Fanuc KAREL source: KT00636.KL

PROGRAM KT00636
%NOLOCKGROUP
VAR
  Y1: ARRAY[2] OF BYTE
  Y2: ARRAY[2] OF BYTE
  OUT: BOOLEAN
BEGIN
  Y1[1] = 2
  Y2[1] = 3
  Y1[1] = 2
  Y2[1] = 3
  OUT = NOT Y1[1]
END KT00636
